PROGRAM MAIN
VAR
	
yellow			: STRING := 'yellow';
blue			: STRING := 'blue';
red				: STRING := 'red';
green 			: STRING := 'green';



END_VAR

END_PROGRAM

(* stored: Version 1.1.0.1
   POU MAIN: Id {c99236d8-b49f-4edf-aac1-911246797e23}, SpecialFunc None *)
